Fanuc KAREL source: KO00150.KL

PROGRAM KO00150
%NOLOCKGROUP
VAR
  R: REAL
  CFG: CONFIG
  OUT: XYZWPR
  N: REAL
BEGIN
  N = 1
  R = 2.0
  CFG.CFG_FLIP = TRUE
  OUT = POS(R, R, R, R, R, N, CFG)
END KO00150
